TYPE ST_VFD_AXIS_REF : FB_VFD_Axis_REF;
END_TYPE

(* stored: Version 1.1.0.1, ProductVersion 3.1.4024.15
   DUT ST_VFD_AXIS_REF: Id {fe227ecc-d6ef-4708-be5c-79c87731157c} *)
